FUNCTION_BLOCK basicEstocagemLodo (* Tanques de estocagem de lodo: sopradores 1+1 com rodizio e intertravamento de nivel das bombas *)
  (* Standard: 61499-2 *)
  (* Version 1.2, 21/10/2026, Hidryco, Hidryco, 1.2: velocidade dos sopradores no automatico (stpVelSopradores em Hz no REQ_PARA, velSO em % no CNF_SO). 1.1: revezamento com horas por soprador (revHabilita, stpTempoB1/B2, padrao do sub-CAT Revezamento) e tempo restante (stsRestanteHor/Min/Seg). 1.0: um soprador sempre ligado no automatico, rodizio por horas (liga o outro antes de desligar), substituicao por indisponibilidade; VA-01/02 e VB-03/04 abertas no automatico; nivel baixo dos tanques com histerese *)
  PACKAGE Hidryco.HidrycoLib;
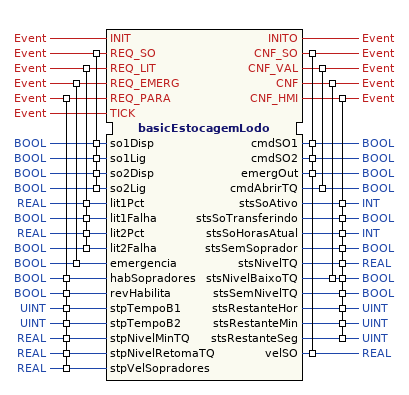
  EVENT_INPUT
    INIT; (* Inicializacao *)
    REQ_SO WITH so1Disp, so1Lig, so2Disp, so2Lig; (* 900-SO-01/02 *)
    REQ_LIT WITH lit1Pct, lit1Falha, lit2Pct, lit2Falha; (* 900-LIT-01/02 (% da faixa) *)
    REQ_EMERG WITH emergencia; (* Emergencia do PCM LODO *)
    REQ_PARA WITH habSopradores, revHabilita, stpTempoB1, stpTempoB2, stpNivelMinTQ, stpNivelRetomaTQ, stpVelSopradores; (* IHM: parametros *)
    TICK; (* Base de tempo de 1 s *)
  END_EVENT
  EVENT_OUTPUT
    INITO; (* Inicializacao concluida *)
    CNF_SO WITH cmdSO1, cmdSO2, emergOut, velSO; (* Comando dos sopradores *)
    CNF_VAL WITH cmdAbrirTQ; (* VA-01, VA-02, VB-03 e VB-04 abertas no automatico *)
    CNF WITH stsNivelBaixoTQ; (* Intertravamento das bombas por nivel dos tanques *)
    CNF_HMI WITH stsSoAtivo, stsSoTransferindo, stsSoHorasAtual, stsSemSoprador, stsNivelTQ, stsNivelBaixoTQ, stsSemNivelTQ, stsRestanteHor, stsRestanteMin, stsRestanteSeg; (* Status para a IHM e alarmes *)
  END_EVENT
  VAR_INPUT
    so1Disp : BOOL; (* SO-01 disponivel para o automatico *)
    so1Lig : BOOL; (* SO-01 ligado *)
    so2Disp : BOOL; (* SO-02 disponivel para o automatico *)
    so2Lig : BOOL; (* SO-02 ligado *)
    lit1Pct : REAL; (* LIT-01 (% da faixa) *)
    lit1Falha : BOOL; (* LIT-01 em falha *)
    lit2Pct : REAL; (* LIT-02 (% da faixa) *)
    lit2Falha : BOOL; (* LIT-02 em falha *)
    emergencia : BOOL; (* Emergencia do PCM LODO *)
    habSopradores : BOOL; (* Sopradores no automatico (um sempre ligado) *)
    revHabilita : BOOL; (* Troca do soprador principal por tempo *)
    stpTempoB1 : UINT; (* Horas do SO-01 como principal; 0 = sem troca por tempo *)
    stpTempoB2 : UINT; (* Horas do SO-02 como principal; 0 = sem troca por tempo *)
    stpNivelMinTQ : REAL; (* Nivel minimo dos tanques para as bombas (%); 0 = sem intertravamento *)
    stpNivelRetomaTQ : REAL; (* Nivel para retomar as bombas (%) *)
    stpVelSopradores : REAL := 60.0; (* Velocidade dos sopradores no automatico (Hz, IHM) *)
  END_VAR
  VAR_OUTPUT
    cmdSO1 : BOOL; (* Liga SO-01 (automatico) *)
    cmdSO2 : BOOL; (* Liga SO-02 (automatico) *)
    emergOut : BOOL; (* Emergencia repassada aos sopradores *)
    cmdAbrirTQ : BOOL; (* Abre VA-01, VA-02, VB-03 e VB-04 (sempre abertas no automatico) *)
    stsSoAtivo : INT; (* Soprador designado: 0 nenhum, 1 SO-01, 2 SO-02 *)
    stsSoTransferindo : BOOL; (* Rodizio em andamento (os dois ligados) *)
    stsSoHorasAtual : INT; (* Horas do soprador atual desde a ultima troca *)
    stsSemSoprador : BOOL; (* Automatico sem nenhum soprador disponivel (risco de sedimentacao) *)
    stsNivelTQ : REAL; (* Nivel usado no intertravamento (maior entre LIT-01 e LIT-02 validos, %) *)
    stsNivelBaixoTQ : BOOL; (* Tanques de estocagem em nivel baixo: bombas suspensas *)
    stsSemNivelTQ : BOOL; (* LIT-01 e LIT-02 em falha: bombas suspensas *)
    stsRestanteHor : UINT; (* Tempo para a troca do soprador principal (h) *)
    stsRestanteMin : UINT; (* Tempo para a troca do soprador principal (min) *)
    stsRestanteSeg : UINT; (* Tempo para a troca do soprador principal (s) *)
    velSO : REAL; (* Referencia dos sopradores no automatico (%, 60 Hz = 100 %) *)
  END_VAR
  VAR
    initDone : BOOL;
    primeiro : BOOL := TRUE;
    ativo : INT;
    tRod : DINT; (* Segundos de operacao do soprador atual *)
    dLim : DINT;
    rest : DINT; (* Segundos ate a troca do soprador principal *)
    rRet : REAL;
    v1 : BOOL;
    v2 : BOOL;
    tVal : INT;
    oldC1 : BOOL;
    oldC2 : BOOL;
    oldEm : BOOL;
    oldBaixo : BOOL;
    sig : INT;
    oldSig : INT := -1;
  END_VAR
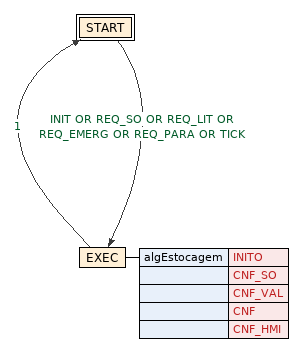
  EC_STATES
    START; (* Estado inicial *)
    EXEC : algEstocagem -> INITO, -> CNF_SO, -> CNF_VAL, -> CNF, -> CNF_HMI; (* Executa a logica; o algoritmo decide quais eventos saem *)
  END_STATES
  EC_TRANSITIONS
    START TO EXEC := INIT OR REQ_SO OR REQ_LIT OR REQ_EMERG OR REQ_PARA OR TICK;
    EXEC TO START := 1;
  END_TRANSITIONS
  ALGORITHM algEstocagem IN ST: (* Logica completa (um unico algoritmo) *)
(* =====================================================================
   basicEstocagemLodo v1.1 - tanques de estocagem de lodo (900, CAT Fase_Solida)
   EF 4.8.1: dois sopradores tri-lobulares 1+1 com rodizio e substituicao;
   em automatico pelo menos um soprador sempre ligado (desligar os dois so em
   manual). VB-03/VB-04 (ar) e VA-01/VA-02 (saida dos tanques) sempre abertas
   no automatico (decisao do usuario). Intertravamento das bombas 900-BO por
   nivel baixo (maior nivel valido entre LIT-01 e LIT-02, % da faixa).
   ===================================================================== *)

INITO   := FALSE;
CNF_SO  := FALSE;
CNF_VAL := FALSE;
CNF     := FALSE;
CNF_HMI := FALSE;

IF INIT THEN
    initDone := TRUE;
    INITO := TRUE;
END_IF;
IF NOT initDone THEN
    RETURN;
END_IF;

(* ---- 1. Sopradores ---- *)
IF NOT habSopradores THEN
    ativo := 0;
    stsSoTransferindo := FALSE;
ELSE
    IF (ativo = 1) AND NOT so1Disp AND so2Disp THEN
        ativo := 2; stsSoTransferindo := FALSE; tRod := 0;          (* substituicao *)
    ELSIF (ativo = 2) AND NOT so2Disp AND so1Disp THEN
        ativo := 1; stsSoTransferindo := FALSE; tRod := 0;
    ELSIF ativo = 0 THEN
        IF so1Disp THEN ativo := 1; tRod := 0;
        ELSIF so2Disp THEN ativo := 2; tRod := 0;
        END_IF;
    END_IF;
    IF ativo = 2 THEN                                               (* horas do soprador atual como principal *)
        dLim := UINT_TO_DINT(stpTempoB2) * 3600;
    ELSE
        dLim := UINT_TO_DINT(stpTempoB1) * 3600;
    END_IF;
    IF NOT stsSoTransferindo AND revHabilita AND (dLim > 0) AND (tRod >= dLim) THEN
        IF ((ativo = 1) AND so2Disp) OR ((ativo = 2) AND so1Disp) THEN
            stsSoTransferindo := TRUE;                              (* liga o outro antes de desligar o atual *)
        END_IF;
    END_IF;
    IF stsSoTransferindo THEN
        IF (ativo = 1) AND so2Lig THEN
            ativo := 2; stsSoTransferindo := FALSE; tRod := 0;
        ELSIF (ativo = 2) AND so1Lig THEN
            ativo := 1; stsSoTransferindo := FALSE; tRod := 0;
        ELSIF ((ativo = 1) AND NOT so2Disp) OR ((ativo = 2) AND NOT so1Disp) THEN
            stsSoTransferindo := FALSE;
        END_IF;
    END_IF;
END_IF;
IF TICK AND (((ativo = 1) AND so1Lig) OR ((ativo = 2) AND so2Lig)) AND (tRod < 2000000000) THEN
    tRod := tRod + 1;
END_IF;
cmdSO1 := habSopradores AND ((ativo = 1) OR (stsSoTransferindo AND (ativo = 2)));
cmdSO2 := habSopradores AND ((ativo = 2) OR (stsSoTransferindo AND (ativo = 1)));
emergOut := emergencia;
velSO := LIMIT(0.0, stpVelSopradores / 0.6, 100.0);   (* IHM em Hz -> % do Motor_Generico *)
stsSoAtivo := ativo;
stsSoHorasAtual := DINT_TO_INT(tRod / 3600);
(* tempo para a troca do principal: 0 = sem troca por tempo (desabilitada, 0 h ou sem soprador) *)
rest := 0;
IF habSopradores AND revHabilita AND (ativo > 0) AND (dLim > 0) AND (tRod < dLim) THEN
    rest := dLim - tRod;
END_IF;
stsRestanteHor := DINT_TO_UINT(rest / 3600);
stsRestanteMin := DINT_TO_UINT((rest MOD 3600) / 60);
stsRestanteSeg := DINT_TO_UINT(rest MOD 60);
stsSemSoprador := habSopradores AND NOT so1Disp AND NOT so2Disp AND NOT so1Lig AND NOT so2Lig;
IF primeiro OR TICK OR (cmdSO1 <> oldC1) OR (cmdSO2 <> oldC2) OR (emergencia <> oldEm) THEN
    CNF_SO := TRUE;
    oldC1 := cmdSO1; oldC2 := cmdSO2; oldEm := emergencia;
END_IF;

(* ---- 2. Valvulas sempre abertas no automatico (reenvio a cada 10 s) ---- *)
cmdAbrirTQ := TRUE;
IF TICK THEN
    tVal := tVal + 1;
END_IF;
IF primeiro OR (tVal >= 10) THEN
    CNF_VAL := TRUE;
    tVal := 0;
END_IF;

(* ---- 3. Nivel dos tanques ---- *)
v1 := NOT lit1Falha;
v2 := NOT lit2Falha;
stsSemNivelTQ := NOT v1 AND NOT v2;
IF v1 AND v2 THEN
    stsNivelTQ := MAX(lit1Pct, lit2Pct);
ELSIF v1 THEN
    stsNivelTQ := lit1Pct;
ELSIF v2 THEN
    stsNivelTQ := lit2Pct;
ELSE
    stsNivelTQ := 0.0;
END_IF;
rRet := MAX(stpNivelRetomaTQ, stpNivelMinTQ);
IF stpNivelMinTQ <= 0.0 THEN
    stsNivelBaixoTQ := FALSE;              (* intertravamento desligado *)
    stsSemNivelTQ := FALSE;
ELSIF stsSemNivelTQ THEN
    stsNivelBaixoTQ := TRUE;               (* sem medicao valida: protege as bombas *)
ELSIF stsNivelTQ < stpNivelMinTQ THEN
    stsNivelBaixoTQ := TRUE;
ELSIF stsNivelTQ >= rRet THEN
    stsNivelBaixoTQ := FALSE;
END_IF;
IF primeiro OR TICK OR (stsNivelBaixoTQ <> oldBaixo) THEN
    CNF := TRUE;
    oldBaixo := stsNivelBaixoTQ;
END_IF;

(* ---- 4. IHM ---- *)
sig := ativo;
IF stsSoTransferindo THEN sig := sig + 4; END_IF;
IF stsSemSoprador THEN sig := sig + 8; END_IF;
IF stsNivelBaixoTQ THEN sig := sig + 16; END_IF;
IF stsSemNivelTQ THEN sig := sig + 32; END_IF;
IF primeiro OR TICK OR REQ_PARA OR (sig <> oldSig) THEN
    CNF_HMI := TRUE;
END_IF;
oldSig := sig;
primeiro := FALSE;
  END_ALGORITHM
END_FUNCTION_BLOCK
